(* PLC project Gaia V8.project, CODESYS CODESYS V3.5 SP22 Patch 2 *)
(* stored: creationDateTime 2026-11-11T09:58:13.2820816, modificationDateTime 2026-11-11T01:17:12.4075064 *)

CONFIGURATION P2_11B
END_CONFIGURATION

CONFIGURATION Module
END_CONFIGURATION

CONFIGURATION Module_3
END_CONFIGURATION

CONFIGURATION Module_1
END_CONFIGURATION

CONFIGURATION Module_2
END_CONFIGURATION

CONFIGURATION <Vide>
END_CONFIGURATION

CONFIGURATION <Vide>
END_CONFIGURATION

CONFIGURATION <Vide>
END_CONFIGURATION

CONFIGURATION <Vide>
END_CONFIGURATION

CONFIGURATION <Vide>
END_CONFIGURATION

CONFIGURATION <Vide>
END_CONFIGURATION

CONFIGURATION <Vide>
END_CONFIGURATION
